(* IEC 61131-3 sources: crb-codesys/retrieval/output/codesys_repo/重型运输系统/modbus/struct, 10 files *)

(* ---- CmdPercentSet.st ---- *)
TYPE CmdPercentSet :
STRUCT
	extendPercent		:WORD;		//0-65535
	retractPercent		:WORD;		//0-65535
END_STRUCT
END_TYPE

(* ---- DeviceUnit.st ---- *)
TYPE DeviceUnit :
STRUCT

	sensor			:SensorInfo;		//传感器参数
	ctrl			:DevPid;			//pid等计算控制执行参数

	vector			:TargetDirect;		//指令运行方向 1-伸出 2-缩回 3-停止
	state			:DevStatus;			//设备状态 0-未知 1-运行 2-伸出到位 3-缩回到位 4-错误

	timeCounter		:INT;				//timeoutCounter超时计数器
	exeCounter		:INT;				//ExecuteCounter额外执行时间计数

	current			:ARRAY[1..2] OF WORD;	//电流mA	[i,j] -> 地轨挡板i的电流，j=1伸出电流，j=2缩回电流

END_STRUCT
END_TYPE

(* ---- DevStatus.st ---- *)
{attribute 'qualified_only'}
{attribute 'strict'}
TYPE DevStatus :
(
	unknown 	:= 0,

	runing		:= 1,

	extended	:= 2,

	retracted	:= 3,

	error		:= 4
);
END_TYPE

(* ---- mdbsRequest.st ---- *)
TYPE mdbsRequest :	//所有请求动作指令数据
STRUCT
	startAddr		:WORD;					//解析起始地址->10
	length			:WORD;					//数据长度/字节->48
	data			:ARRAY[10..57] OF WORD;	//指令数据

	arrNew		:ARRAY [1..4,0..15] OF BOOL;
	arrLast		:ARRAY [1..4,0..15] OF BOOL;

END_STRUCT
END_TYPE

(* ---- mdbsResponse.st ---- *)
TYPE mdbsResponse :	//所有响应状态数据回送
STRUCT
	startAddr		:WORD;							//解析起始地址->110
	length			:WORD;							//字节长度->210

	data			:ARRAY[110..319] OF WORD;		//位置数据

END_STRUCT
END_TYPE

(* ---- mdbsStruct.st ---- *)
TYPE mdbsStruct :
STRUCT
	request		:mdbsRequest;				//请求动作指令
	response	:mdbsResponse;			//响应动作指令-天地轨所有

END_STRUCT
END_TYPE

(* ---- SensorInfo.st ---- *)
TYPE SensorInfo :
STRUCT

	position	:REAL;	//实时位移
	speed		:REAL;	//实时速度

	//记录最大最小位移值
	retractVal	:REAL;	//缩回到位值
	extendVal	:REAL;	//伸出到位值

END_STRUCT
END_TYPE

(* ---- TargetDirect.st ---- *)
{attribute 'qualified_only'}
{attribute 'strict'}
TYPE TargetDirect :
(
	extend 	:= 1,	//伸出

	retract := 2,	//缩回

	stop	:= 3	//停止
);
END_TYPE

(* ---- UIMode.st ---- *)
TYPE UIMode :
STRUCT
	manualButtonSet			:BOOL;		//手动复位按钮模式
	usePID					:BOOL;		//使用pid
	autoEnable				:BOOL;		//自动使能
	manualPercentSet		:BOOL;		//手动设定比例量
	manualSetPid			:BOOL;		//手动调节pid参数，可通过pid测试界面设定目标位移值

	syncExt					:BOOL;		//同步伸
	syncRct					:BOOL;		//同步缩

	hydPowerOn				:BOOL;		//液压站开启 modbus 使用
	hydPowerOff				:BOOL;		//液压站关闭 modbus 使用
	hydPowerReset			:BOOL;
END_STRUCT
END_TYPE

(* ---- UIUnit.st ---- *)
TYPE UIUnit :
STRUCT
	//cmd
	pwrEnable			:BOOL;		//比例阀使能   power-enable
	pwrPercent			:REAL;		//比例阀百分比 power-percent 0-100

	//button
	btnExtend			:BOOL;
	btnRetract			:BOOL;
	btnStop				:BOOL;
	btnLast				:TargetDirect;	//上次动作方向

	//info display
	name				:STRING;	//挡板名
	wname				:WSTRING;	//山河命名
	hzname				:WSTRING;	//hua zhong ming ming
	postion				:REAL;		//位移值
	speed				:REAL;
	extendPercent		:REAL;		//伸出百分比 extend-percent

END_STRUCT
END_TYPE
